// TIA Portal V21 export
// export: Created 2026-11-10T07:35:16.5073805Z, ExportSetting WithDefaults, DisplayName Totally Integrated Automation Portal, DisplayVersion V21 Update 3, DisplayName STEP 7 Professional, DisplayVersion V21 Update 3, DisplayName STEP 7 Safety, DisplayVersion V21, DisplayName Tech WebApplication, DisplayVersion V21, DisplayName WinCC Basic/Comfort/Advanced, DisplayVersion V21 Update 3, DisplayName WinCC Unified, DisplayVersion V21 Update 3
FUNCTION_BLOCK "FB_Lad_ex125"   // FB47, LAD
{ S7_Optimized_Access := 'TRUE' }
VERSION : 0.1
// stored: AutoNumber true, IsIECCheckEnabled false, IsRetainMemResEnabled false, MemoryReserve 100, SetENOAutomatically false, UDAEnableTagReadback false
   VAR_INPUT
      v_mode : UInt;
      v_ob : OB_ANY;
      v_ret_val : Int;
   END_VAR
   VAR_IN_OUT
      v_info : Variant;
   END_VAR
BEGIN

REGION Network 1: RT_INFO - Read out runtime statistics
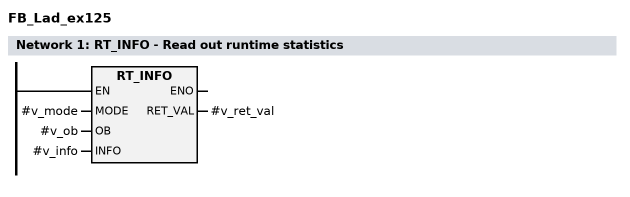
   RUNG wire#powerrail
      RT_INFO(MODE := #v_mode, OB := #v_ob, Ret_Val => #v_ret_val, INFO := #v_info)
   END_RUNG
   // the same network as SCL:
   #v_ret_val := RT_INFO(MODE := #v_mode, OB := #v_ob, INFO := #v_info);
END_REGION
END_FUNCTION_BLOCK
